KUKA KRL program: folge11.src, folge11.dat

--- folge11.src ---
&ACCESS RVP
&REL 1
&COMMENT bt2krl vw-ks24 production Folge 11 plan 16#A1BE
DEF FOLGE11()
   ; Generated by bt2krl 0.1.0 from bt2plc plan bt_1792156523_scene_fit (cell scene_fit), PLAN_ID 16#A1BE
   ; Robot robot2 (R2), controller robot2, model unknown, joint mapping identity
   ; Profile vw-ks24 (VW KS24 / TPVW 8.1.8).
   ; Do not edit: regenerate with bt2krl (plain KRL, no inline forms).
   ; Production Folge: 3 ops; per op: op index BT_PKTNR, interlock request + MAKRO20 handshake, motion (exact stop at the end), hold, interlock release
   ; The VW tech package does the Folge handshake (cell.src, AUE_INIT/WAIT/END).
   ;FOLD AUE INIT
      VW(#VW_AUE_INIT,TRUE)
      PENTER:
      INTERRUPT DECL 10 WHEN $CYCFLAG[254]==FALSE DO VW(#FB_STOP,TRUE)
      INTERRUPT ON 10
      INT10=TRUE
   ;ENDFOLD
   ;FOLD VWP0 P0 10 PCT
      ; P0 = home: VW_INIT runs BAS(#INITMOV); AUE_WAIT later sets $H_POS here
      VW(#VW_INIT,TRUE)
      VW_USR_R (#USR_INIT)
      BAS(#VEL_PTP,10)
      $APO.CPTP=100
      PTP P0
      $OUT[15]=TRUE ; PF0 Grundstellung
      ; MAKRO0 RUECKSETZEN_EA: resets A33-A96 (also the tool releases)
      SEL_RES=SELECT(#MAKRO,0,TRUE,,,,,FALSE)
   ;ENDFOLD
   ;FOLD VWAUEWAIT
      VW(#VW_AUE_WAIT,TRUE )
      IF N_VW==TRUE THEN
         GOTO PEXIT
      ENDIF
   ;ENDFOLD
   ;FOLD VWSTART 16#00000003
      ; release every interlock this robot uses: IL01=V1 IL02=V2
      $OUT[15]=FALSE ; PF0 off
      ; MAKRO50 Ini Merker: the cyclic flags of the driving conditions
      SEL_RES=SELECT(#MAKRO,50,TRUE,,,,,FALSE)
      $OUT[41]=TRUE ; release V1
      $OUT[42]=TRUE ; release V2
   ;ENDFOLD
   ;FOLD VWFB 16#00000000
      VALCYCFL30=$CYCFLAG[254]
      $CYCFLAG[254]=($CYCFLAG[30]) AND $CYCFLAG[255] OR ($TIMER[61]<0)
      VW(#FB_CHECK,TRUE)
   ;ENDFOLD
   ;FOLD OP 1 W01 MASK 16#00000002
      ; zones IL02
      BT_PKTNR=1
      ;FOLD VWLOCK 16#00000002
         ; enter IL02=V2
         $OUT[82]=TRUE ; request V2
         ; MAKRO20 semantics, inline for these interlocks only
         $OUT[42]=$OUT[42] OR $OUT[82]
         ; PLC grant of the request
         $LOOP_MSG[]="E82"
         $LOOP_CONT=TRUE
         WAIT FOR ($IN[82]) OR (NOT $LOOP_CONT AND ($MODE_OP<>#EX))
         $LOOP_MSG[]="                                                                                                                                "
         ; partner release
         $LOOP_MSG[]="E42"
         $LOOP_CONT=TRUE
         WAIT FOR ($IN[42]) OR (NOT $LOOP_CONT AND ($MODE_OP<>#EX))
         $LOOP_MSG[]="                                                                                                                                "
         $OUT[42]=FALSE ; occupied
         $OUT[82]=FALSE
      ;ENDFOLD
      ;FOLD VWFB 16#00000002
         VALCYCFL30=$CYCFLAG[254]
         $CYCFLAG[254]=($CYCFLAG[30] AND $IN[42]) AND $CYCFLAG[255] OR ($TIMER[61]<0)
         VW(#FB_CHECK,TRUE)
      ;ENDFOLD
      BAS(#VEL_PTP,2)
      PTP P1 C_PTP
      BAS(#VEL_PTP,3)
      PTP P2 C_PTP
      BAS(#VEL_PTP,5)
      PTP P3 C_PTP
      BAS(#VEL_PTP,7)
      PTP P4 C_PTP
      BAS(#VEL_PTP,8)
      PTP P5 C_PTP
      BAS(#VEL_PTP,9)
      PTP P6 C_PTP
      BAS(#VEL_PTP,11)
      PTP P7 C_PTP
      BAS(#VEL_PTP,10)
      PTP P8 C_PTP
      BAS(#VEL_PTP,9)
      PTP P9 C_PTP
      BAS(#VEL_PTP,7)
      PTP P10 C_PTP
      BAS(#VEL_PTP,6)
      PTP P11 C_PTP
      BAS(#VEL_PTP,4)
      PTP P12 C_PTP
      BAS(#VEL_PTP,3)
      PTP P13 C_PTP
      BAS(#VEL_PTP,2)
      PTP P14 C_PTP
      BAS(#VEL_PTP,6)
      PTP P15 C_PTP
      BAS(#VEL_PTP,8)
      PTP P16 C_PTP
      BAS(#VEL_PTP,3)
      PTP P17
      WAIT SEC 0.5 ; hold
      ;FOLD VWUNLOCK 16#00000002
         ; leave IL02=V2
         $OUT[42]=TRUE ; release V2
      ;ENDFOLD
      ;FOLD VWFB 16#00000000
         VALCYCFL30=$CYCFLAG[254]
         $CYCFLAG[254]=($CYCFLAG[30]) AND $CYCFLAG[255] OR ($TIMER[61]<0)
         VW(#FB_CHECK,TRUE)
      ;ENDFOLD
      WAIT SEC 0.1 ; step dwell
   ;ENDFOLD
   ;FOLD OP 2 W03 MASK 16#00000001
      ; zones IL01
      BT_PKTNR=2
      ;FOLD VWLOCK 16#00000001
         ; enter IL01=V1
         $OUT[81]=TRUE ; request V1
         ; MAKRO20 semantics, inline for these interlocks only
         $OUT[41]=$OUT[41] OR $OUT[81]
         ; PLC grant of the request
         $LOOP_MSG[]="E81"
         $LOOP_CONT=TRUE
         WAIT FOR ($IN[81]) OR (NOT $LOOP_CONT AND ($MODE_OP<>#EX))
         $LOOP_MSG[]="                                                                                                                                "
         ; partner release
         $LOOP_MSG[]="E41"
         $LOOP_CONT=TRUE
         WAIT FOR ($IN[41]) OR (NOT $LOOP_CONT AND ($MODE_OP<>#EX))
         $LOOP_MSG[]="                                                                                                                                "
         $OUT[41]=FALSE ; occupied
         $OUT[81]=FALSE
      ;ENDFOLD
      ;FOLD VWFB 16#00000001
         VALCYCFL30=$CYCFLAG[254]
         $CYCFLAG[254]=($CYCFLAG[30] AND $IN[41]) AND $CYCFLAG[255] OR ($TIMER[61]<0)
         VW(#FB_CHECK,TRUE)
      ;ENDFOLD
      BAS(#VEL_PTP,4)
      PTP P18 C_PTP
      PTP P19 C_PTP
      BAS(#VEL_PTP,10)
      PTP P20 C_PTP
      BAS(#VEL_PTP,13)
      PTP P21 C_PTP
      BAS(#VEL_PTP,11)
      PTP P22 C_PTP
      BAS(#VEL_PTP,7)
      PTP P23 C_PTP
      BAS(#VEL_PTP,3)
      PTP P24 C_PTP
      BAS(#VEL_PTP,6)
      PTP P25 C_PTP
      BAS(#VEL_PTP,8)
      PTP P26 C_PTP
      BAS(#VEL_PTP,3)
      PTP P27
      WAIT SEC 0.5 ; hold
      ;FOLD VWUNLOCK 16#00000001
         ; leave IL01=V1
         $OUT[41]=TRUE ; release V1
      ;ENDFOLD
      ;FOLD VWFB 16#00000000
         VALCYCFL30=$CYCFLAG[254]
         $CYCFLAG[254]=($CYCFLAG[30]) AND $CYCFLAG[255] OR ($TIMER[61]<0)
         VW(#FB_CHECK,TRUE)
      ;ENDFOLD
      WAIT SEC 0.1 ; step dwell
   ;ENDFOLD
   ;FOLD OP 3 HOME MASK 16#00000002
      ; zones IL02
      BT_PKTNR=3
      ;FOLD VWLOCK 16#00000002
         ; enter IL02=V2
         $OUT[82]=TRUE ; request V2
         ; MAKRO20 semantics, inline for these interlocks only
         $OUT[42]=$OUT[42] OR $OUT[82]
         ; PLC grant of the request
         $LOOP_MSG[]="E82"
         $LOOP_CONT=TRUE
         WAIT FOR ($IN[82]) OR (NOT $LOOP_CONT AND ($MODE_OP<>#EX))
         $LOOP_MSG[]="                                                                                                                                "
         ; partner release
         $LOOP_MSG[]="E42"
         $LOOP_CONT=TRUE
         WAIT FOR ($IN[42]) OR (NOT $LOOP_CONT AND ($MODE_OP<>#EX))
         $LOOP_MSG[]="                                                                                                                                "
         $OUT[42]=FALSE ; occupied
         $OUT[82]=FALSE
      ;ENDFOLD
      ;FOLD VWFB 16#00000002
         VALCYCFL30=$CYCFLAG[254]
         $CYCFLAG[254]=($CYCFLAG[30] AND $IN[42]) AND $CYCFLAG[255] OR ($TIMER[61]<0)
         VW(#FB_CHECK,TRUE)
      ;ENDFOLD
      BAS(#VEL_PTP,5)
      PTP P28 C_PTP
      BAS(#VEL_PTP,2)
      PTP P29 C_PTP
      BAS(#VEL_PTP,5)
      PTP P30 C_PTP
      BAS(#VEL_PTP,8)
      PTP P31 C_PTP
      BAS(#VEL_PTP,10)
      PTP P32 C_PTP
      BAS(#VEL_PTP,12)
      PTP P33 C_PTP
      BAS(#VEL_PTP,14)
      PTP P34 C_PTP
      PTP P35 C_PTP
      BAS(#VEL_PTP,13)
      PTP P36 C_PTP
      BAS(#VEL_PTP,12)
      PTP P37 C_PTP
      BAS(#VEL_PTP,10)
      PTP P38 C_PTP
      BAS(#VEL_PTP,8)
      PTP P39 C_PTP
      BAS(#VEL_PTP,5)
      PTP P40 C_PTP
      BAS(#VEL_PTP,2)
      PTP P41
      ;FOLD VWMAKRO 15
         ; Gesamtfertigmeldung
         SEL_RES=SELECT(#MAKRO,15,TRUE,,,,,FALSE)
      ;ENDFOLD
      ;FOLD VWUNLOCK 16#00000002
         ; leave IL02=V2
         $OUT[42]=TRUE ; release V2
      ;ENDFOLD
      ;FOLD VWFB 16#00000000
         VALCYCFL30=$CYCFLAG[254]
         $CYCFLAG[254]=($CYCFLAG[30]) AND $CYCFLAG[255] OR ($TIMER[61]<0)
         VW(#FB_CHECK,TRUE)
      ;ENDFOLD
      WAIT SEC 0.1 ; step dwell
   ;ENDFOLD
   BT_PKTNR=0
   ;FOLD AUE END
      VW(#VW_AUE_END,TRUE)
      GOTO PENTER
      PEXIT:
   ;ENDFOLD
END

--- folge11.dat ---
&ACCESS RVP
&REL 1
&COMMENT bt2krl vw-ks24 data Folge 11 plan 16#A1BE
DEFDAT FOLGE11
   ; Generated by bt2krl 0.1.0 from bt2plc plan bt_1792156523_scene_fit (cell scene_fit), PLAN_ID 16#A1BE
   ; Robot robot2 (R2), controller robot2, model unknown, joint mapping identity
   ; Profile vw-ks24 (VW KS24 / TPVW 8.1.8).
   ; Do not edit: regenerate with bt2krl (plain KRL, no inline forms).
   EXT BAS (BAS_COMMAND :IN,REAL :IN )
   ; interface to the VW standard routines (as every VW Folge .dat declares them)
   EXT VW (VW_COMMAND :IN,BOOL :IN,REAL :IN,REAL :IN,REAL :IN,REAL :IN,BOOL :IN,E6POS :IN )
   EXT VW_USR_R (VW_USER_CMD :IN,INT :IN,REAL :IN,REAL :IN,REAL :IN,REAL :IN,REAL :IN,REAL :IN,BOOL :IN )
   EXTFCT INT SELECT (SUBTYPE :IN,INT :IN,BOOL :IN,ARI_TYP :IN,INT :IN,BOOL_TYP :IN,INT :IN,BOOL :IN)
   DECL AXIS P0={A1 45.0,A2 -90.0,A3 90.0,A4 0.0,A5 0.0,A6 0.0}
   DECL AXIS P1={A1 44.7829,A2 -89.9274,A3 90.0007,A4 0.0,A5 0.5792,A6 -1.1959}
   DECL AXIS P2={A1 44.1614,A2 -89.7195,A3 90.0027,A4 0.0,A5 2.2369,A6 -4.6186}
   DECL AXIS P3={A1 43.1805,A2 -89.3915,A3 90.0058,A4 0.0,A5 4.8532,A6 -10.0208}
   DECL AXIS P4={A1 41.8851,A2 -88.9583,A3 90.01,A4 0.0,A5 8.3083,A6 -17.1549}
   DECL AXIS P5={A1 39.4506,A2 -88.1442,A3 90.0178,A4 0.0,A5 14.8017,A6 -30.5623}
   DECL AXIS P6={A1 36.5613,A2 -87.178,A3 90.0271,A4 0.0,A5 22.5083,A6 -46.475}
   DECL AXIS P7={A1 24.5256,A2 -83.153,A3 90.0658,A4 0.0,A5 54.6107,A6 -112.7595}
   DECL AXIS P8={A1 21.5184,A2 -82.1473,A3 90.0755,A4 0.0,A5 62.6319,A6 -129.3216}
   DECL AXIS P9={A1 19.7288,A2 -81.5489,A3 90.0812,A4 0.0,A5 67.4051,A6 -139.1775}
   DECL AXIS P10={A1 17.4796,A2 -80.7967,A3 90.0885,A4 0.0,A5 73.4042,A6 -151.5643}
   DECL AXIS P11={A1 16.3359,A2 -80.4142,A3 90.0921,A4 0.0,A5 76.4549,A6 -157.8633}
   DECL AXIS P12={A1 15.5291,A2 -80.1444,A3 90.0947,A4 0.0,A5 78.6069,A6 -162.3067}
   DECL AXIS P13={A1 15.2661,A2 -80.0565,A3 90.0956,A4 0.0,A5 79.3084,A6 -163.7552}
   DECL AXIS P14={A1 15.0489,A2 -79.9839,A3 90.0963,A4 0.0,A5 79.8876,A6 -164.9511}
   DECL AXIS P15={A1 15.0489,A2 -79.8382,A3 90.6698,A4 0.0,A5 79.1684,A6 -164.9511}
   DECL AXIS P16={A1 15.0489,A2 -79.6225,A3 91.5053,A4 0.0,A5 78.1172,A6 -164.9511}
   DECL AXIS P17={A1 15.0489,A2 -78.7572,A3 94.1833,A4 0.0,A5 74.5738,A6 -164.9511}
   DECL AXIS P18={A1 15.0298,A2 -79.8762,A3 90.5449,A4 0.0,A5 79.3313,A6 -164.9702}
   DECL AXIS P19={A1 13.7592,A2 -79.9905,A3 90.0976,A4 0.0,A5 79.8929,A6 -166.2408}
   DECL AXIS P20={A1 9.2892,A2 -80.0151,A3 90.0809,A4 0.0,A5 79.9342,A6 -170.7108}
   DECL AXIS P21={A1 -8.1126,A2 -80.0749,A3 90.1766,A4 0.0,A5 79.8983,A6 -188.1126}
   DECL AXIS P22={A1 -11.544,A2 -80.0849,A3 90.2027,A4 0.0,A5 79.8822,A6 -191.544}
   DECL AXIS P23={A1 -13.8724,A2 -80.0914,A3 90.2214,A4 0.0,A5 79.87,A6 -193.8724}
   DECL AXIS P24={A1 -14.7302,A2 -80.0938,A3 90.2286,A4 0.0,A5 79.8652,A6 -194.7302}
   DECL AXIS P25={A1 -14.7302,A2 -79.9478,A3 90.8022,A4 0.0,A5 79.1457,A6 -194.7302}
   DECL AXIS P26={A1 -14.7302,A2 -79.7318,A3 91.6378,A4 0.0,A5 78.094,A6 -194.7302}
   DECL AXIS P27={A1 -14.7302,A2 -78.865,A3 94.3164,A4 0.0,A5 74.5486,A6 -194.7302}
   DECL AXIS P28={A1 -14.7302,A2 -79.9187,A3 90.9391,A4 0.0,A5 78.9797,A6 -194.7302}
   DECL AXIS P29={A1 -14.0312,A2 -80.0367,A3 90.9281,A4 0.0,A5 78.0554,A6 -192.4514}
   DECL AXIS P30={A1 -12.0585,A2 -80.3697,A3 90.8971,A4 0.0,A5 75.4469,A6 -186.0199}
   DECL AXIS P31={A1 -8.9984,A2 -80.8861,A3 90.849,A4 0.0,A5 71.4007,A6 -176.0436}
   DECL AXIS P32={A1 -5.0374,A2 -81.5547,A3 90.7867,A4 0.0,A5 66.1631,A6 -163.1301}
   DECL AXIS P33={A1 1.3232,A2 -82.6282,A3 90.6867,A4 0.0,A5 57.7527,A6 -142.3935}
   DECL AXIS P34={A1 8.5122,A2 -83.8416,A3 90.5737,A4 0.0,A5 48.2468,A6 -118.9561}
   DECL AXIS P35={A1 25.428,A2 -86.6966,A3 90.3077,A4 0.0,A5 25.8795,A6 -63.8078}
   DECL AXIS P36={A1 30.6317,A2 -87.5749,A3 90.2259,A4 0.0,A5 18.9988,A6 -46.8431}
   DECL AXIS P37={A1 35.3072,A2 -88.364,A3 90.1524,A4 0.0,A5 12.8165,A6 -31.6001}
   DECL AXIS P38={A1 39.2682,A2 -89.0326,A3 90.0901,A4 0.0,A5 7.579,A6 -18.6866}
   DECL AXIS P39={A1 42.3283,A2 -89.5491,A3 90.042,A4 0.0,A5 3.5328,A6 -8.7103}
   DECL AXIS P40={A1 44.301,A2 -89.882,A3 90.011,A4 0.0,A5 0.9243,A6 -2.2789}
   DECL AXIS P41={A1 45.0,A2 -90.0,A3 90.0,A4 0.0,A5 0.0,A6 0.0}
ENDDAT
